// TIA Portal V19 export
TYPE "ST_Home"
   STRUCT
      Execute : Bool;
      Busy : Bool;
      Done : Bool;
      Error : Bool;
      ErrorID : Word;
      CommandAborted : Bool;
      Mode : Int;
      Position : Int;
      ReferencePosition : Real;
   END_STRUCT;
END_TYPE
